Fanuc KAREL source: KC00013.KL

PROGRAM KC00013
%NOLOCKGROUP
%ENVIRONMENT PBQMGR
VAR
  I: INTEGER
  J: INTEGER
  K: INTEGER
  R: REAL
  B: BOOLEAN
  S: STRING[80]
  T: STRING[80]
  P: PATH
  Q: PATH
  QT: QUEUE_TYPE
  AI: ARRAY[8] OF INTEGER
  AB: ARRAY[244] OF BYTE
BEGIN
  GET_QUEUE(QT,AI,I,J,K)
END KC00013
